Fanuc KAREL source: KE00003.KL

PROGRAM KE00003
%NOLOCKGROUP
%ENVIRONMENT REGOPE
VAR
  I: INTEGER
  S: STRING[80]
  STATUS: INTEGER
BEGIN
  I = 1
  S = 'TEST'
  SET_PREG_CMT(I, S, STATUS)
END KE00003
